(* IEC 61131-3 sources: Caravan/Archiv/12-04-19/Stations/MachineControl/MachineControl/Class/Timer_Class, 1 file *)

(* ---- Timer_Class.st ---- *)
(*!
<Class
	Name               = "Timer_Class"
	Revision           = "0.0"
	RealtimeTask       = "false"
	CyclicTask         = "true"
	DefCyclictime      = "100 µs"
	BackgroundTask     = "false"
	Sigmatek           = "false"
	OSInterface        = "false"
	HighPriority       = "false"
	Automatic          = "false"
	UpdateMode         = "Prescan"
	SharedCommandTable = "true"
	Objectsize         = "(630,180)">
	<Channels>
		<Server Name="ClassSvr" Visualized="false" Remotely="true" Initialize="false" WriteProtected="true" Retentive="false"/>
		<Server Name="Nachtmodus_S" Visualized="true" Remotely="true" Initialize="false" WriteProtected="false" Retentive="SRam"/>
	</Channels>
</Class>
*)
Timer_Class : CLASS
  //Servers:
	ClassSvr 	: SvrChCmd_DINT;
	Nachtmodus_S 	: SvrCh_DINT;
  //Clients:
  //Variables:
  //Functions:

	FUNCTION VIRTUAL GLOBAL CyWork
		VAR_INPUT
			EAX 	: UDINT;
		END_VAR
		VAR_OUTPUT
			state (EAX) 	: UDINT;
		END_VAR;
  //Tables:
	FUNCTION @STD
		VAR_OUTPUT
			ret_code	: CONFSTATES;
		END_VAR;
	FUNCTION GLOBAL TAB @CT_;
END_CLASS;

FUNCTION VIRTUAL GLOBAL Timer_Class::CyWork
	VAR_INPUT
		EAX 	: UDINT;
	END_VAR
	VAR_OUTPUT
		state (EAX) 	: UDINT;
	END_VAR

	state := READY;

END_FUNCTION
